(* IEC 61131-3 sources: Versio-VersionControlSystem/fixtures/projects/TC3_PlcSample_reStrText/TC3_PlcSample_reStrText/LibraryDocumentationSample Project/LibPOUs/B_DocuElements/Text blocks, 3 files *)

(* ---- FB_Libdoc_BlockQuote.st ---- *)
(*
This is a top-level paragraph.

    This paragraph belongs to a first-level block quote.

    This is the second paragraph of the first-level block quote.

        This paragraph belongs to a second-level block quote.

Another top-level paragraph.

        This paragraph belongs to a second-level block quote.

    This paragraph belongs to a first-level block quote. The
    second-level block quote above is inside this first-level
    block quote.
*)

FUNCTION_BLOCK FB_Libdoc_BlockQuote
VAR_INPUT
    nVarA : INT;
    nVarB : INT;
END_VAR
VAR_OUTPUT
    nSum : INT;
END_VAR
VAR
END_VAR

(* ---- FB_Libdoc_LineBlock.st ---- *)
(*
Line blocks are useful where the structure of lines is significant.

| Each new line begins with
| a vertical bar ("|").
|     Line breaks and initial indents
|     are preserved.
| Continuation lines are wrapped
  portions of long lines; they begin
  with spaces in place of vertical bars.

    | Each new line begins with
    | a vertical bar ("|").
    |     Line breaks and initial indents
    |     are preserved.
    | Continuation lines are wrapped
      portions of long lines; they begin
      with spaces in place of vertical bars.
*)

FUNCTION_BLOCK FB_Libdoc_LineBlock
VAR_INPUT
    nVarA : INT;
    nVarB : INT;
END_VAR
VAR_OUTPUT
    nSum : INT;
END_VAR
VAR
END_VAR

(* ---- FB_Libdoc_Paragraph.st ---- *)
(*
This is a paragraph.

Paragraphs line up at their left edges, and are normally separated
by blank lines.
*)

FUNCTION_BLOCK FB_Libdoc_Paragraph
VAR_INPUT
    nVarA : INT;
    nVarB : INT;
END_VAR
VAR_OUTPUT
    nSum : INT;
END_VAR
VAR
END_VAR
